Fanuc KAREL source: KD00035.KL

PROGRAM KD00035
%NOLOCKGROUP
VAR
  I: INTEGER
  J: INTEGER
  B: BOOLEAN
  R: REAL
  S: STRING[80]
BEGIN
  CONDITION[1]:
  WHEN DIN[1] = ON DO
    CONTINUE
  ENDCONDITION
END KD00035
